(* IEC 61131-3 sources: plc_generation_empirical_study/datasets/_archive/pre_native_plcverif_20260810/tasks/C07_E01_linear_scaling/negative_control, 1 file *)

(* ---- NC1.st ---- *)
FUNCTION_BLOCK C07_E01_linear_scaling
VAR_INPUT
    Raw : INT;
END_VAR
VAR_OUTPUT
    Engineering : REAL;
END_VAR

Engineering := INT_TO_REAL(Raw) * 0.2;

END_FUNCTION_BLOCK
